Fanuc KAREL source: KA00093.KL

PROGRAM KA00093
%NOLOCKGROUP
VAR
  SRC: JOINTPOS
  DST: VECTOR
BEGIN
  DST = SRC
END KA00093
